INTERFACE I_DriveAxis

METHOD Execute
END_METHOD

METHOD Enable
END_METHOD

METHOD Disable
END_METHOD

METHOD SetVelocity
VAR_INPUT
	velocityInMPerS : LREAL;
END_VAR
END_METHOD

METHOD TryReset : BOOL
END_METHOD

PROPERTY PositionInM : LREAL
GET
END_GET
END_PROPERTY

PROPERTY VelocityInMPerS : LREAL
GET
END_GET
END_PROPERTY

PROPERTY IsReady : BOOL
GET
END_GET
END_PROPERTY

PROPERTY Error : HardwareError
GET
END_GET
END_PROPERTY

END_INTERFACE

(* stored: Version 1.1.0.1, ProductVersion 3.1.4026.12
   Itf I_DriveAxis: Id {10aea2a4-a0f9-52d9-bfb9-5a25b6bff0c4}
   Method Execute: Id {1e83eb23-3ac7-570f-8c9f-0f9d28ced79d}
   Method Enable: Id {0d90f66d-ffe8-5589-b620-609e5c982203}
   Method Disable: Id {b4433f01-4685-5393-961d-f2156ab8ac26}
   Method SetVelocity: Id {ebdf5207-0d77-5272-8477-dc32725f3a2f}
   Method TryReset: Id {7ddb3653-ef36-558c-b73c-97250a736f88}
   Property PositionInM: Id {3ebba2b9-13aa-5538-b04e-af7dfe5b536c}
   Get Get: Id {17e4dc54-f244-5f17-99c1-082aa86e65e0}
   Property VelocityInMPerS: Id {802943f5-1cd8-55bf-8544-e49974164e4a}
   Get Get: Id {97ec4d4b-bb1f-5de2-96b8-ccf6bbbfa3b1}
   Property IsReady: Id {a55d4ba7-b37d-5808-9a32-c19d01fe0749}
   Get Get: Id {0d0031f4-9b45-5338-ae22-86c8d88e7c49}
   Property Error: Id {077314a0-d591-5246-a87a-d40cbf37e8c3}
   Get Get: Id {2c10dc1c-882a-5ba7-b59b-9e30c87023ed} *)
